(* PLC project Simulatie Sorteer Station, CODESYS CODESYS V3.5 SP16 Patch 7, author Rene Potters/Gerard Harkema *)
(* stored: creationDateTime 2026-11-26T15:39:48.4972208, version 0.1.0, modificationDateTime 2026-11-26T15:37:02.1644744, organization Avans *)
(* Simulatie voor opstelling Sorteer Station. *)

VAR_GLOBAL  (* GVL *)
  Ix_Resetknop : BOOL;  (* Indrukken resetknop *)
  Ix_Hand : BOOL;  (* Keuzeknop staat op hand *)
  Ix_Auto : BOOL;  (* Keuzeknop staat op auto *)
  Ix_Noodstop : BOOL;  (* Indrukken noodstop *)
  Ix_MagazijnLeeg : BOOL;  (* Bekers magazijn zijn op *)
  Ix_UitstoterBekerIn : BOOL;  (* Beker is uit dekselmagazijn gestoten *)
  Ix_UitstoterBekerUit : BOOL;  (* Uitstoter Beker haalt nieuwe beker op *)
  Ix_Stopknop : BOOL := TRUE;  (* Indrukken startknop *)
  Ix_Startknop : BOOL;  (* Indrukken stopknop *)
  Ix_PersluchtAanwezig : BOOL;  (* Perslucht is aanwezig *)
  Ix_VacuumAanwezig : BOOL;  (* Werkstuk door overzetter opgepakt *)
  Ix_OverzetterIsLinks : BOOL;  (* Overzetter haalt beker op(linker pos.) *)
  Ix_OverzetterIsRechts : BOOL;  (* Overzetter plaatst beker op afgifteplaats *)
  Qx_BekerUitstoten : BOOL;  (* Beker uit magazijn stoten *)
  Qx_VacuumAan : BOOL;  (* Beker oppakken *)
  Qx_BekerLossen : BOOL;  (* Beker loslaten *)
  Qx_OverzetterLinks : BOOL;  (* Overzetter naar bekermagazijn *)
  Qx_OverzetterRechts : BOOL;  (* Overzetter naar afgifteplaats *)
  Qx_GeleLamp : BOOL;  (* Visualisatie invisible Gele vlak *)
  Qx_GroeneLamp : BOOL;  (* Visualisatie invisible groene vlak *)
  Qx_RodeLamp : BOOL;  (* Visualisatie invisible rode vlak *)
END_VAR

CONFIGURATION Device
  RESOURCE ApplicationSt ON PLC
    TASK MainTask(INTERVAL := T#20ms, PRIORITY := 1);
    TASK Simulatie(INTERVAL := T#20ms, PRIORITY := 1);
    PROGRAM Main WITH MainTask : Main;
    PROGRAM MagazijnSim WITH Simulatie : MagazijnSim;
    PROGRAM OverzetterSim WITH Simulatie : OverzetterSim;
  END_RESOURCE
END_CONFIGURATION

CONFIGURATION Basic
END_CONFIGURATION

CONFIGURATION <Empty>
END_CONFIGURATION

CONFIGURATION <Empty>
END_CONFIGURATION

CONFIGURATION <Empty>
END_CONFIGURATION

CONFIGURATION <Empty>
END_CONFIGURATION

CONFIGURATION <Empty>
END_CONFIGURATION

CONFIGURATION <Empty>
END_CONFIGURATION

CONFIGURATION <Empty>
END_CONFIGURATION

CONFIGURATION <Empty>
END_CONFIGURATION

CONFIGURATION <Empty>
END_CONFIGURATION

CONFIGURATION <Empty>
END_CONFIGURATION

CONFIGURATION <Empty>
END_CONFIGURATION
